(* IEC 61131-3 sources: avi-aoi-management/scripts/ai-eval/ngau-nhien/kho/st-ud9-ghi-dich-loai-bo/mau/src, 2 files *)

(* ---- LoaiBoAOI.st ---- *)
FUNCTION_BLOCK LoaiBoAOI
VAR_INPUT
    ENCODER : BOOL;
    CO_SAN_PHAM : BOOL;
    LOI_AOI : BOOL;
    RESET : BOOL;
    VI_TRI_GAT : INT;
    T_GAT : TIME;
END_VAR
VAR_OUTPUT
    CAN_GAT : BOOL;
    DEM_GAT : DINT;
    SO_O_LOI : INT;
END_VAR
VAR
    rtEnc : R_TRIG;
    tg : ThanhGhiDich;
    xungGat : TP;
    toi : BOOL;
END_VAR
    rtEnc(CLK := ENCODER);
    tg(DICH := rtEnc.Q AND NOT RESET, GHI := CO_SAN_PHAM AND LOI_AOI AND NOT RESET, XOA := RESET, VI_TRI := VI_TRI_GAT);
    (* sản phẩm lỗi vừa được dịch tới vị trí gạt *)
    toi := rtEnc.Q AND NOT RESET AND VI_TRI_GAT >= 1 AND VI_TRI_GAT <= 32 AND tg.Q;
    IF RESET THEN
        DEM_GAT := 0;
    ELSIF toi THEN
        DEM_GAT := DEM_GAT + 1;
    END_IF
    xungGat(IN := toi, PT := T_GAT);
    CAN_GAT := xungGat.Q;
    SO_O_LOI := tg.SO_O;
END_FUNCTION_BLOCK

(* ---- ThanhGhiDich.st ---- *)
FUNCTION_BLOCK ThanhGhiDich
VAR_INPUT
    DICH : BOOL;
    GHI : BOOL;
    XOA : BOOL;
    VI_TRI : INT;
END_VAR
VAR_OUTPUT
    Q : BOOL;
    SO_O : INT;
END_VAR
VAR
    o : ARRAY[0..32] OF BOOL;
    i : INT;
END_VAR
    IF XOA THEN
        FOR i := 0 TO 32 DO o[i] := FALSE; END_FOR
    ELSE
        IF DICH THEN
            FOR i := 32 TO 1 BY -1 DO o[i] := o[i - 1]; END_FOR
            o[0] := FALSE;
        END_IF
        IF GHI THEN
            o[0] := TRUE;
        END_IF
    END_IF
    IF VI_TRI >= 0 AND VI_TRI <= 32 THEN
        Q := o[VI_TRI];
    ELSE
        Q := FALSE;
    END_IF
    SO_O := 0;
    FOR i := 0 TO 32 DO
        IF o[i] THEN SO_O := SO_O + 1; END_IF
    END_FOR
END_FUNCTION_BLOCK
